Fanuc KAREL source: kt00911.KL

-- PROVISIONAL review KL for V770-1; original PC SHA256 51d15b072f169ae6c4bba862c18a3eb6c38a16364859ceecf709fe7af157235a
-- Incomplete behavior may be omitted. Consult companion uncertainty JSON. Do not deploy.
PROGRAM KT00911
%NOLOCKGROUP
BEGIN
  -- UNRESOLVED_PC offsets 5-31; opcodes 27,27,49,7E,AD,31,4A
  -- UNRESOLVED_PC offsets 36-40; opcodes 7F
END KT00911
